FUNCTION_BLOCK HMI_BLOCKS (* Composite Function Block Type *)
  (* Standard: 61499-2 *)
  (* Version 0.0, 3/6/2020, jhunjhp1, nxtControl GmbH, template *)
  PACKAGE Main;
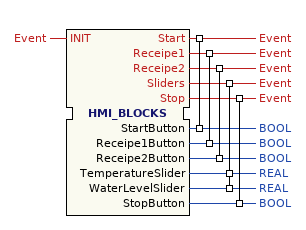
  EVENT_INPUT
    INIT; (* Initialization Request *)
  END_EVENT
  EVENT_OUTPUT
    Start WITH StartButton; (* Initialization Confirm *)
    Receipe1 WITH Receipe1Button; (* Execution Confirmation *)
    Receipe2 WITH Receipe2Button;
    Sliders WITH TemperatureSlider, WaterLevelSlider;
    Stop WITH StopButton;
  END_EVENT
  VAR_OUTPUT
    StartButton : BOOL; (* Output event qualifier *)
    Receipe1Button : BOOL;
    Receipe2Button : BOOL;
    TemperatureSlider : REAL;
    WaterLevelSlider : REAL;
    StopButton : BOOL;
  END_VAR
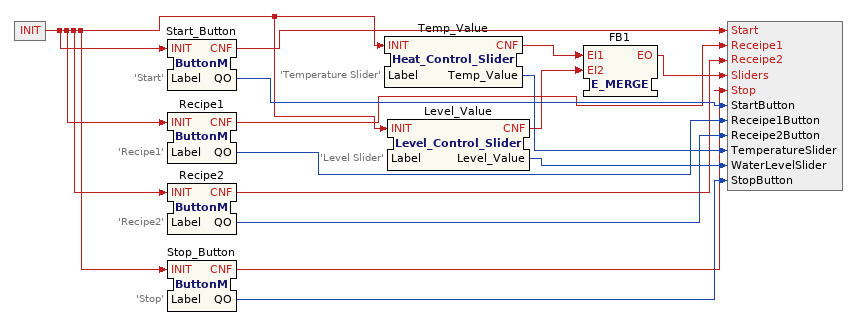
  FBS
    Start_Button : ButtonM(Label := 'Start');
    Temp_Value : Heat_Control_Slider(Label := 'Temperature Slider');
    Level_Value : Level_Control_Slider(Label := 'Level Slider');
    Recipe1 : ButtonM(Label := 'Recipe1');
    Recipe2 : ButtonM(Label := 'Recipe2');
    Stop_Button : ButtonM(Label := 'Stop');
    FB1 : E_MERGE;
  END_FBS
  EVENT_CONNECTIONS
    INIT TO Start_Button.INIT;
    INIT TO Recipe1.INIT;
    INIT TO Recipe2.INIT;
    INIT TO Stop_Button.INIT;
    Start_Button.CNF TO Start;
    Recipe1.CNF TO Receipe1;
    Recipe2.CNF TO Receipe2;
    Stop_Button.CNF TO Stop;
    Temp_Value.CNF TO FB1.EI1;
    Level_Value.CNF TO FB1.EI2;
    FB1.EO TO Sliders;
    INIT TO Temp_Value.INIT;
    INIT TO Level_Value.INIT;
  END_CONNECTIONS
  DATA_CONNECTIONS
    Start_Button.QO TO StartButton;
    Temp_Value.Temp_Value TO TemperatureSlider;
    Level_Value.Level_Value TO WaterLevelSlider;
    Recipe1.QO TO Receipe1Button;
    Recipe2.QO TO Receipe2Button;
    Stop_Button.QO TO StopButton;
  END_CONNECTIONS
END_FUNCTION_BLOCK
